(* IEC 61131-3 sources: llm-plc-st-eval/data/definitivo/gpt-4o-2024-08-06/A3/zero_shot, 3 files *)

(* ---- ejec_1.st ---- *)
```pascal
FUNCTION_BLOCK FB_Com
VAR
    // Entradas
    txReq : BOOL;
    rxOk : BOOL;
    rxData : INT;

    // Salidas
    txData : INT;
    ocupado : BOOL;
    ok : BOOL;
    error : BOOL;
    nIntentos : INT;

    // Variables internas
    txReqPrev : BOOL; // Para detectar flancos
    intentoActual : INT; // Contador de intentos
    timer : TON; // Temporizador para los 500 ms
    intentoExitoso : BOOL; // Indica si el intento fue exitoso
END_VAR

// Inicialización de variables
IF NOT ocupado THEN
    txData := 100; // Valor de prueba
    intentoActual := 0;
    intentoExitoso := FALSE;
    ok := FALSE;
    error := FALSE;
END_IF

// Detección de flanco ascendente en txReq
IF txReq AND NOT txReqPrev THEN
    IF NOT ocupado THEN
        // Iniciar nuevo intercambio
        ocupado := TRUE;
        intentoActual := 1;
        nIntentos := intentoActual;
        timer(IN := TRUE, PT := T#500MS);
    END_IF
END_IF

// Guardar estado anterior de txReq
txReqPrev := txReq;

// Lógica de intercambio
IF ocupado THEN
    // Verificar si el temporizador ha expirado
    timer(IN := TRUE);
    IF timer.Q THEN
        // Intento fallido, incrementar contador de intentos
        intentoActual := intentoActual + 1;
        IF intentoActual > 3 THEN
            // Todos los intentos fallaron
            error := TRUE;
            ocupado := FALSE;
        ELSE
            // Iniciar nuevo intento
            nIntentos := intentoActual;
            timer(IN := TRUE, PT := T#500MS);
        END_IF
    ELSE
        // Verificar si el intento es exitoso
        IF rxOk AND (rxData = txData) THEN
            intentoExitoso := TRUE;
            ok := TRUE;
            ocupado := FALSE;
        END_IF
    END_IF
END_IF
```

Este código implementa un intercambio de petición/respuesta con un dispositivo externo, manejando hasta 3 intentos y verificando el éxito de cada intento dentro de un plazo de 500 milisegundos.

(* ---- ejec_2.st ---- *)
```pascal
FUNCTION_BLOCK FB_Com
VAR
    // Entradas
    txReq : BOOL;
    rxOk : BOOL;
    rxData : INT;

    // Salidas
    txData : INT := 0;
    ocupado : BOOL := FALSE;
    ok : BOOL := FALSE;
    error : BOOL := FALSE;
    nIntentos : INT := 0;

    // Variables internas
    intentoActual : INT := 0;
    tiempoInicio : TIME;
    tiempoActual : TIME;
    esperandoRespuesta : BOOL := FALSE;
    valorPrueba : INT := 100;
END_VAR

// Código del bloque de función
IF NOT ocupado AND txReq THEN
    // Iniciar nuevo intercambio
    txData := valorPrueba;
    ocupado := TRUE;
    ok := FALSE;
    error := FALSE;
    intentoActual := 1;
    nIntentos := intentoActual;
    tiempoInicio := TIME(); // Captura el tiempo actual
    esperandoRespuesta := TRUE;
ELSIF ocupado THEN
    // Si estamos ocupados, verificar el estado del intento actual
    tiempoActual := TIME();

    IF esperandoRespuesta THEN
        // Verificar si se recibió respuesta correcta
        IF rxOk AND rxData = valorPrueba THEN
            // Respuesta correcta
            ok := TRUE;
            ocupado := FALSE;
            esperandoRespuesta := FALSE;
        ELSIF (tiempoActual - tiempoInicio) >= T#500MS THEN
            // Tiempo de espera agotado, intentar de nuevo
            intentoActual := intentoActual + 1;
            IF intentoActual > 3 THEN
                // Todos los intentos fallaron
                error := TRUE;
                ocupado := FALSE;
                esperandoRespuesta := FALSE;
            ELSE
                // Iniciar nuevo intento
                nIntentos := intentoActual;
                tiempoInicio := tiempoActual; // Reiniciar tiempo de inicio
            END_IF
        END_IF
    END_IF
END_IF
```

Este código implementa un intercambio de petición/respuesta con un dispositivo externo, manejando hasta 3 intentos y verificando la respuesta dentro de un plazo de 500 ms.

(* ---- ejec_3.st ---- *)
```pascal
FUNCTION_BLOCK FB_Com
VAR
    // Entradas
    txReq: BOOL;
    rxOk: BOOL;
    rxData: INT;

    // Salidas
    txData: INT;
    ocupado: BOOL;
    ok: BOOL;
    error: BOOL;
    nIntentos: INT;

    // Variables internas
    intentoActual: INT := 0;
    tiempoInicio: TIME;
    tiempoTranscurrido: TIME;
    txReqPrev: BOOL := FALSE;
    intentoExitoso: BOOL := FALSE;
END_VAR

VAR CONSTANT
    VALOR_PRUEBA: INT := 100;
    TIEMPO_MAXIMO: TIME := T#500MS;
    MAX_INTENTOS: INT := 3;
END_VAR

// Lógica del bloque de funciones
IF NOT ocupado THEN
    // Detectar flanco ascendente de txReq
    IF txReq AND NOT txReqPrev THEN
        // Iniciar un nuevo intercambio
        txData := VALOR_PRUEBA;
        ocupado := TRUE;
        ok := FALSE;
        error := FALSE;
        intentoActual := 1;
        nIntentos := intentoActual;
        tiempoInicio := TIME(); // Guardar el tiempo de inicio
    END_IF;
ELSE
    // Intercambio en curso
    tiempoTranscurrido := TIME() - tiempoInicio;

    IF rxOk AND (rxData = VALOR_PRUEBA) THEN
        // Intento exitoso
        intentoExitoso := TRUE;
        ok := TRUE;
        ocupado := FALSE;
    ELSIF tiempoTranscurrido >= TIEMPO_MAXIMO THEN
        // Intento fallido, verificar si hay más intentos
        intentoActual := intentoActual + 1;
        IF intentoActual > MAX_INTENTOS THEN
            // Todos los intentos fallaron
            error := TRUE;
            ocupado := FALSE;
        ELSE
            // Iniciar un nuevo intento
            nIntentos := intentoActual;
            tiempoInicio := TIME(); // Reiniciar el tiempo de inicio
        END_IF;
    END_IF;
END_IF;

// Actualizar txReqPrev para detectar flancos
txReqPrev := txReq;
```

Este código implementa un intercambio de petición/respuesta con un dispositivo externo, manejando hasta 3 intentos y verificando el eco del valor transmitido.
